(* PLC project Vn_chain_deep, Beckhoff Automation GmbH TwinCAT PLC Control 3.5.13.21 *)
(* stored: creationDateTime 1970-01-01T00:00:00 *)

PROGRAM Vn_chain_deep

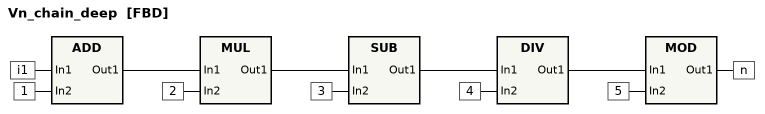
(* FBD diagram, written out as Structured Text *)
n := ((i1 + 1) * 2 - 3) / 4 MOD 5;
END_PROGRAM
